(* CODESYS project station.library
   DefaultNamespace: KOSTAL.AF2024.Core.Station
   DocFormat: reStructuredText
   Description: contain base Framework for station-internal connection
   Author: Frank Dümpelmann
   Title: KOSTAL.AF2024.Core.Station
   Version: 1.0.0.0
   Company: KOSTAL GmbH & Co.KG
   Placeholder: KOSTAL.AF2024.Core.Station

Project tree, tasks and I/O mapping:
  libraries: KOSTAL.AF2024.Core.FileLogger, 1.0.0.0 (KOSTAL GmbH & Co.KG); KOSTAL.AF2024.Core.ID, 1.0.0.0 (KOSTAL GmbH & Co.KG); KOSTAL.AF2024.Core.MainControl, 1.0.0.0 (KOSTAL GmbH & Co.KG); KOSTAL.AF2024.Core.Process, 1.0.0.0 (KOSTAL GmbH & Co.KG); KOSTAL.AF2024.Core.Settings, 1.0.0.0 (KOSTAL GmbH & Co.KG); KOSTAL.AF2024.Core.StringTools, 1.0.0.0 (KOSTAL GmbH & Co.KG); KOSTAL.AF2024.Core.System, 1.0.0.0 (KOSTAL GmbH & Co.KG); KOSTAL.AF2024.Core.Text, 1.0.0.0 (KOSTAL GmbH & Co.KG)
  1_Station_Free/
    function block FB_Station_Free [ST]: _getNameAndID, _ID_TO_WSTRING, _log, _log_isReady, _parameterControl, _TextReader, FB_init, linkLogger, LogText, Condition, Condition_Owner, ID, Message, Message_Owner, Name, TextPath
    interface I_Station_Free: Condition, ID, Message, Name
    interface I_Station_Free_Owner: Condition, Condition_Owner, ID, LogText, Message, Message_Owner, Name
  2_Station_Controlled/
    function block FB_Station_Controlled [ST]: _log, MainControl, State, State_Owner, Step, Step_Owner
    interface I_Station_Controlled: MainControl, State, Step
    interface I_Station_Controlled_Owner: MainControl, State, State_Owner, Step, Step_Owner
  Project Information/
    function F_GetCompany [ST]
    function F_GetTitle [ST]
    function F_GetVersion [ST]
  Version/
    global variables Global_Version
*)

// Version/Global_Version
{attribute 'TcGenerated'}
{attribute 'no-analysis'}
{attribute 'linkalways'}
// This function has been automatically generated from the project information.
VAR_GLOBAL CONSTANT
	{attribute 'const_non_replaced'}
	stLibVersion_KOSTAL_AF2024_Core_Station : ST_LibVersion := (iMajor := 1, iMinor := 0, iBuild := 0, iRevision := 0, nFlags := 0, sVersion := '1.0.0.0');
END_VAR

// 1_Station_Free/FB_Station_Free
FUNCTION_BLOCK PUBLIC FB_Station_Free IMPLEMENTS I_Station_Free, I_Station_Free_Owner

VAR
	//=============================================================================================================================================================
	//=============================================================================================================================================================
	_ID	: KOSTAL_AF2024_Core_ID.T_ID;

	//=======================================================================================================================================
	_Name	: KOSTAL_AF2024_Core_Settings.T_MaxString;	//localized name of station

	_condition			: KOSTAL_AF2024_Core_Process.FB_processCondition;

	_Logger	: KOSTAL_AF2024_Core_FileLogger.I_Logger;
	
	//=============================================================================================================================================================
	_message				: KOSTAL_AF2024_Core_Process.T_messageText_3_lines;
	//=============================================================================================================================================================

	//Text
	_TextPath		: KOSTAL_AF2024_Core_Settings.T_MaxString_UTF8;
	_Text			: KOSTAL_AF2024_Core_Text.FB_Handler_Slave;	//local text content
	
	_TextInitialized	: BOOL;
END_VAR

METHOD PROTECTED _getNameAndID : KOSTAL_AF2024_Core_Settings.T_MaxString

VAR
	_c	: KOSTAL_AF2024_Core_StringTools.FB_Concat;
END_VAR


_c.Clear();
_c.addContent(_Name);
_c.addContent("[");
_c.addContent(_ID.name);
_c.addContent("(");
_c.addContent(DINT_TO_WSTRING(_ID.key));
_c.addContent(")");
_c.addContent("]");
_getNameAndID:= _c.getResult();
_c.Clear();
END_METHOD

METHOD PROTECTED _ID_TO_WSTRING : KOSTAL_AF2024_Core_Settings.T_MaxString

VAR
	_c	: KOSTAL_AF2024_Core_StringTools.FB_Concat;
END_VAR


_c.Clear();
_c.addContent(_ID.name);
_c.addContent("(");
_c.addContent(DINT_TO_WSTRING(_ID.key));
_c.addContent(")");
_ID_TO_WSTRING:= _c.getResult();
_c.Clear();
END_METHOD

METHOD PROTECTED _log : BOOL
VAR_INPUT
	Text	: KOSTAL_AF2024_Core_Settings.T_MaxString;
END_VAR

IF _Logger = 0 THEN 
	RETURN;	
END_IF
IF NOT _Logger.State.success THEN 
	RETURN;	
END_IF

_Logger.ID					:= _ID_TO_WSTRING();
_Logger.name				:= _Name;


_Logger.addLine(Text);

_log:= TRUE;
END_METHOD

METHOD PROTECTED _log_isReady : BOOL

IF _Logger = 0 							THEN RETURN;	END_IF
IF NOT _Logger.State.success	THEN RETURN;	END_IF

_log_isReady:= TRUE;
END_METHOD

(*
	| Add here your implementation of Interface controls like:

	| IF _IgetTime = 0 THEN

	| 	_message.clear();

	| 	_textHandlerCommon.clearVars();
	| 	_message.line_01:= 'Parameter Fail';
	| 	_message.line_02:= 'Interface _IgetTime is not linked';

	| 	_condition.setMessage(4999, _message);

	| ELSE
	
	| 	_parameterControl:= TRUE;

	| END_IF
*)

METHOD PROTECTED _parameterControl : BOOL
VAR_INPUT
END_VAR

// no parameters to control in base
_parameterControl:= TRUE;

(* Add here your implementation of Interface controls like:

_parameterControl:= FALSE;

IF _IgetTime = 0 THEN

	_message.clear();

	_textHandlerCommon.clearVars();
	_message.line_01:= 'Parameter Fail';
	_message.line_02:= 'Interface _IgetTime is not linked';

	_condition.setMessage(4999, _message);

ELSE
	
	_parameterControl:= TRUE;

END_IF
*)
END_METHOD

//Returns true if text was initialized once
METHOD PROTECTED _TextReader : BOOL;
VAR_INPUT
END_VAR

_Text.Path:= _TextPath;
_Text.FBmain();

IF _text.State.fail THEN
	_message.clear();	
	_message.line_01:= "TextHandler";
	_message.line_02:= _Text.State.description;
	_condition.setMessage(_condition.PriorityLevel_Error, _message);
ELSIF NOT _Text.Valid THEN
	_name := _ID.name;
	_message.clear();	
	_message.line_01:= "TextHandler";
	_message.line_02:= _Text.State.description;
	_condition.setMessage(_condition.PriorityLevel_MasterMessage + 999, _message);//Overwrite all other messages
END_IF


IF _text.LoadedLanguage <> '' THEN
	_textInitialized := TRUE;
END_IF
_TextReader := _textInitialized;
END_METHOD

METHOD FB_init : BOOL
VAR_INPUT
	bInitRetains 	: BOOL; // if TRUE, the retain variables are initialized (warm start / cold start)
	bInCopyCode 	: BOOL;  // if TRUE, the instance afterwards gets moved into the copy code (online change)
	ID_Name				: KOSTAL_AF2024_Core_Settings.T_MaxString;
	ID_Key				: DINT;
	CommonText		: KOSTAL_AF2024_Core_Text.I_Text;
END_VAR

_ID.name:= ID_Name;
_ID.key	:= ID_Key;

_text.linkCommonText(CommonText);
END_METHOD

METHOD PUBLIC linkLogger
VAR_INPUT
	logger	: KOSTAL_AF2024_Core_FileLogger.I_Logger;
END_VAR

_Logger:= logger;
END_METHOD

(*
	These PUBLIC methods are required to make the log function usable for interface participants (such as cylinders).
*)
METHOD PUBLIC LogText : BOOL
VAR_INPUT
	Text	: KOSTAL_AF2024_Core_Settings.T_MaxString;
END_VAR
LogText:= _log(Text);
END_METHOD

PROPERTY PUBLIC Condition : KOSTAL_AF2024_Core_Process.I_processCondition
GET

Condition := _condition;
END_GET
END_PROPERTY

PROPERTY PUBLIC Condition_Owner : KOSTAL_AF2024_Core_Process.I_processCondition_Owner
GET

Condition_Owner := _condition;
END_GET
END_PROPERTY

PROPERTY PUBLIC ID : KOSTAL_AF2024_Core_ID.I_T_ID
GET

ID := _ID;
END_GET
END_PROPERTY

PROPERTY PUBLIC Message : KOSTAL_AF2024_Core_Process.I_T_messageText_3_lines
GET

Message := _message;
END_GET
END_PROPERTY

PROPERTY PUBLIC Message_Owner : KOSTAL_AF2024_Core_Process.I_T_messageText_3_lines_Owner
GET

Message_Owner := _message;
END_GET
END_PROPERTY

//localized name of station
PROPERTY PUBLIC Name : KOSTAL_AF2024_Core_Settings.T_MaxString
GET

Name:= _Name;
END_GET
SET

_Name:= Name;
END_SET
END_PROPERTY

PROPERTY PUBLIC TextPath : KOSTAL_AF2024_Core_Settings.T_MaxString_UTF8
GET

TextPath:= _TextPath;
END_GET
SET

_TextPath:= TextPath;
END_SET
END_PROPERTY

END_FUNCTION_BLOCK

// 1_Station_Free/I_Station_Free
INTERFACE I_Station_Free EXTENDS KOSTAL_AF2024_Core_System.I_Interface

PROPERTY PUBLIC Condition : KOSTAL_AF2024_Core_Process.I_processCondition
GET
END_GET
END_PROPERTY

PROPERTY PUBLIC ID : KOSTAL_AF2024_Core_ID.I_T_ID
GET
END_GET
END_PROPERTY

PROPERTY PUBLIC Message : KOSTAL_AF2024_Core_Process.I_T_messageText_3_lines
GET
END_GET
END_PROPERTY

//localized name of station
PROPERTY PUBLIC Name : KOSTAL_AF2024_Core_Settings.T_MaxString
GET
END_GET
END_PROPERTY

END_INTERFACE

// 1_Station_Free/I_Station_Free_Owner
INTERFACE I_Station_Free_Owner EXTENDS KOSTAL_AF2024_Core_System.I_Interface

PROPERTY PUBLIC Condition : KOSTAL_AF2024_Core_Process.I_processCondition
GET
END_GET
END_PROPERTY

PROPERTY PUBLIC Condition_Owner : KOSTAL_AF2024_Core_Process.I_processCondition_Owner
GET
END_GET
END_PROPERTY

PROPERTY PUBLIC ID : KOSTAL_AF2024_Core_ID.I_T_ID
GET
END_GET
END_PROPERTY

(*
	These PUBLIC methods are required to make the log function usable for interface participants (such as cylinders).
*)
METHOD PUBLIC LogText : BOOL
VAR_INPUT
	Text	: KOSTAL_AF2024_Core_Settings.T_MaxString;
END_VAR
END_METHOD

PROPERTY PUBLIC Message : KOSTAL_AF2024_Core_Process.I_T_messageText_3_lines
GET
END_GET
END_PROPERTY

PROPERTY PUBLIC Message_Owner : KOSTAL_AF2024_Core_Process.I_T_messageText_3_lines_Owner
GET
END_GET
END_PROPERTY

//localized name of station
PROPERTY PUBLIC Name : KOSTAL_AF2024_Core_Settings.T_MaxString
GET
END_GET
SET
END_SET
END_PROPERTY

END_INTERFACE

// 2_Station_Controlled/FB_Station_Controlled
(*
	Extend the FB_FR_Station class with conectivity to a main control 
*)
FUNCTION_BLOCK PUBLIC FB_Station_Controlled EXTENDS FB_Station_Free IMPLEMENTS I_Station_Controlled, I_Station_Controlled_Owner
VAR
	_step		: KOSTAL_AF2024_Core_Process.FB_ProcessStep_Control;
	_state		: KOSTAL_AF2024_Core_MainControl.T_ParticipantState;

	_mainControl		: KOSTAL_AF2024_Core_MainControl.FB_Participant(ID:= _ID, Condition:= _condition, State:= _state);
END_VAR

METHOD PROTECTED _log : BOOL
VAR_INPUT
	Text	: KOSTAL_AF2024_Core_Settings.T_MaxString;
END_VAR
IF _Logger = 0 THEN 
	RETURN;	
END_IF


_Logger.stepNumber	:= _step.actual;



_log:= SUPER^._log(Text);
END_METHOD

PROPERTY MainControl : KOSTAL_AF2024_Core_MainControl.I_Participant
GET

MainControl:= _mainControl;
END_GET
END_PROPERTY

PROPERTY PUBLIC State : KOSTAL_AF2024_Core_MainControl.I_T_participantState; //KOSTAL_AF2024_Core_process.FB_plcState;
GET


State := _state;
END_GET
END_PROPERTY

PROPERTY PUBLIC State_Owner : KOSTAL_AF2024_Core_MainControl.I_T_participantState_Owner; //KOSTAL_AF2024_Core_process.FB_plcState;
GET


State_Owner := _state;
END_GET
END_PROPERTY

PROPERTY PUBLIC Step : KOSTAL_AF2024_Core_Process.I_ProcessStep_Control
GET
Step := _step;
END_GET
END_PROPERTY

PROPERTY PUBLIC Step_Owner : KOSTAL_AF2024_Core_Process.I_ProcessStep_Control_Owner
GET
Step_Owner := _step;
END_GET
END_PROPERTY

END_FUNCTION_BLOCK

// 2_Station_Controlled/I_Station_Controlled
INTERFACE I_Station_Controlled EXTENDS I_Station_Free

PROPERTY PUBLIC MainControl : KOSTAL_AF2024_Core_MainControl.I_Participant
GET
END_GET
END_PROPERTY

PROPERTY PUBLIC State : KOSTAL_AF2024_Core_MainControl.I_T_participantState; //KOSTAL_AF2024_Core_process.FB_plcState;
GET
END_GET
END_PROPERTY

PROPERTY PUBLIC Step : KOSTAL_AF2024_Core_Process.I_ProcessStep_Control
GET
END_GET
END_PROPERTY

END_INTERFACE

// 2_Station_Controlled/I_Station_Controlled_Owner
INTERFACE I_Station_Controlled_Owner EXTENDS I_Station_Free_Owner

PROPERTY PUBLIC MainControl : KOSTAL_AF2024_Core_MainControl.I_Participant
GET
END_GET
END_PROPERTY

PROPERTY PUBLIC State : KOSTAL_AF2024_Core_MainControl.I_T_participantState; //KOSTAL_AF2024_Core_process.FB_plcState;
GET
END_GET
END_PROPERTY

PROPERTY PUBLIC State_Owner : KOSTAL_AF2024_Core_MainControl.I_T_participantState_Owner; //KOSTAL_AF2024_Core_process.FB_plcState;
GET
END_GET
END_PROPERTY

PROPERTY PUBLIC Step : KOSTAL_AF2024_Core_Process.I_ProcessStep_Control
GET
END_GET
END_PROPERTY

PROPERTY PUBLIC Step_Owner : KOSTAL_AF2024_Core_Process.I_ProcessStep_Control_Owner
GET
END_GET
END_PROPERTY

END_INTERFACE

// Project Information/F_GetCompany
// This function has been automatically generated from the project information.
{attribute 'signature_flag' := '1073741824'}
{attribute 'TcGenerated'}
{attribute 'no-analysis'}
FUNCTION F_GetCompany : WSTRING
VAR_INPUT
	
END_VAR

F_GetCompany := "KOSTAL GmbH & Co.KG";

END_FUNCTION

// Project Information/F_GetTitle
// This function has been automatically generated from the project information.
{attribute 'signature_flag' := '1073741824'}
{attribute 'TcGenerated'}
{attribute 'no-analysis'}
FUNCTION F_GetTitle : WSTRING
VAR_INPUT
	
END_VAR

F_GetTitle := "KOSTAL.AF2024.Core.Station";

END_FUNCTION

// Project Information/F_GetVersion
// This function has been automatically generated from the project information.
{attribute 'signature_flag' := '1073741824'}
{attribute 'TcGenerated'}
{attribute 'no-analysis'}
FUNCTION F_GetVersion : ST_LibVersion
VAR_INPUT
	
END_VAR

F_GetVersion.iMajor := 1;
F_GetVersion.iMinor := 0;
F_GetVersion.iBuild := 0;
F_GetVersion.iRevision := 0;
F_GetVersion.sVersion := '1.0.0.0';
F_GetVersion.nFlags := 0;

END_FUNCTION
